(* IEC 61131-3 sources: rusty/tests/lit/multi/duplicate_unit_ctor_basename_1723, 1 file *)

(* ---- main.st ---- *)
FUNCTION main : DINT
    main := g_in_a + g_in_b;
    IF main = 33 THEN
        printf('ok$N');
    END_IF;
END_FUNCTION
